// TIA Portal project "kelishangliao" (V15)

(* hardware
DEVICE "S7300/ET200M station_1"  S7-300 station
   slot 0: "导轨_0"  Rail  6ES7 390-1***0-0AA0
   slot 2: "PLC_1"  CPU 314C-2 PN/DP  6ES7 314-6EH04-0AB0  V3.3
      slot 2: "PROFINET 接口_1"  PN-IO
         slot 1: "Port_1"  Port
         slot 2: "Port_2"  Port
      slot 5: "DI 24/DO 16_1"  DI24/DO16
      slot 6: "AI 5/AO 2_1"  AI5/AO2
      slot 7: "计数_1"  Counter
      slot 8: "定位_1"  Positioning
*)

// ===== PLC "PLC_1"  CPU 314C-2 PN/DP =====

VAR_GLOBAL   // PLC tag table "默认变量表"
   "开始按钮" AT %I0.0 : Bool;
   "复位按钮" AT %I0.1 : Bool;
   "停止按钮" AT %I0.4 : Bool;
   "上电" AT %I0.5 : Bool;
   "空瓶到位" AT %I1.0 : Bool;
   "夹瓶处电眼" AT %I1.1 : Bool;
   "颗粒有无" AT %I1.2 : Bool;
   "末端颗粒到位" AT %I1.5 : Bool;
   "主传输带" AT %Q0.0 : Bool;
   "颗粒料传送带" AT %Q0.1 : Bool;
   "旋转气缸" AT %Q0.2 : Bool;
   "升降气缸" AT %Q0.3 : Bool;
   "夹瓶气缸" AT %Q0.4 : Bool;
   "推料颗粒气缸" AT %Q0.5 : Bool;
   "吸盘_电磁阀" AT %Q0.7 : Bool;
   "空瓶输送带_变频器" AT %Q1.0 : Bool;
   "开始灯_绿" AT %Q1.6 : Bool;
   "复位灯_橙" AT %Q1.7 : Bool;
   "M0" AT %M10.0 : Bool;
   "M1" AT %M10.1 : Bool;
   "M2" AT %M10.2 : Bool;
   "M3" AT %M10.3 : Bool;
   "M4" AT %M10.4 : Bool;
   "M5" AT %M10.5 : Bool;
   "M6" AT %M10.6 : Bool;
   "M7" AT %M10.7 : Bool;
   "Tag_1" AT %MD100 : Time;
   "Tag_2" AT %MD104 : Time;
   "Tag_3" AT %MD108 : Time;
   "Tag_4" AT %MD112 : Time;
   "Tag_5" AT %MD116 : Time;
   "Tag_6" AT %MD120 : Time;
   "Tag_7" AT %MD124 : Time;
   "Tag_8" AT %MD128 : Time;
   "Tag_9" AT %MD132 : Time;
   "Tag_10" AT %MW200 : Int;
END_VAR

ORGANIZATION_BLOCK "Main"   // OB1, LAD
TITLE = "Main Program Sweep (Cycle)"
{ S7_Optimized_Access := 'FALSE' }
VERSION : 0.1
   VAR_TEMP
      OB1_EV_CLASS : Byte;   // Bits 0-3 = 1 (Coming event), Bits 4-7 = 1 (Event class 1)
      OB1_SCAN_1 : Byte;   // 1 (Cold restart scan 1 of OB 1), 3 (Scan 2-n of OB 1)
      OB1_PRIORITY : Byte;   // Priority of OB Execution
      OB1_OB_NUMBR : Byte;   // 1 (Organization block 1, OB1)
      OB1_RESERVED_1 : Byte;   // Reserved for system
      OB1_RESERVED_2 : Byte;   // Reserved for system
      OB1_PREV_CYCLE : Int;   // Cycle time of previous OB1 scan (milliseconds)
      OB1_MIN_CYCLE : Int;   // Minimum cycle time of OB1 (milliseconds)
      OB1_MAX_CYCLE : Int;   // Maximum cycle time of OB1 (milliseconds)
      OB1_DATE_TIME : Date_And_Time;   // Date and time OB1 started
   END_VAR
   VAR_TEMP   // added for the SCL form of the ladder/FBD networks
      _w1 : Bool;
   END_VAR
BEGIN

REGION Network 1
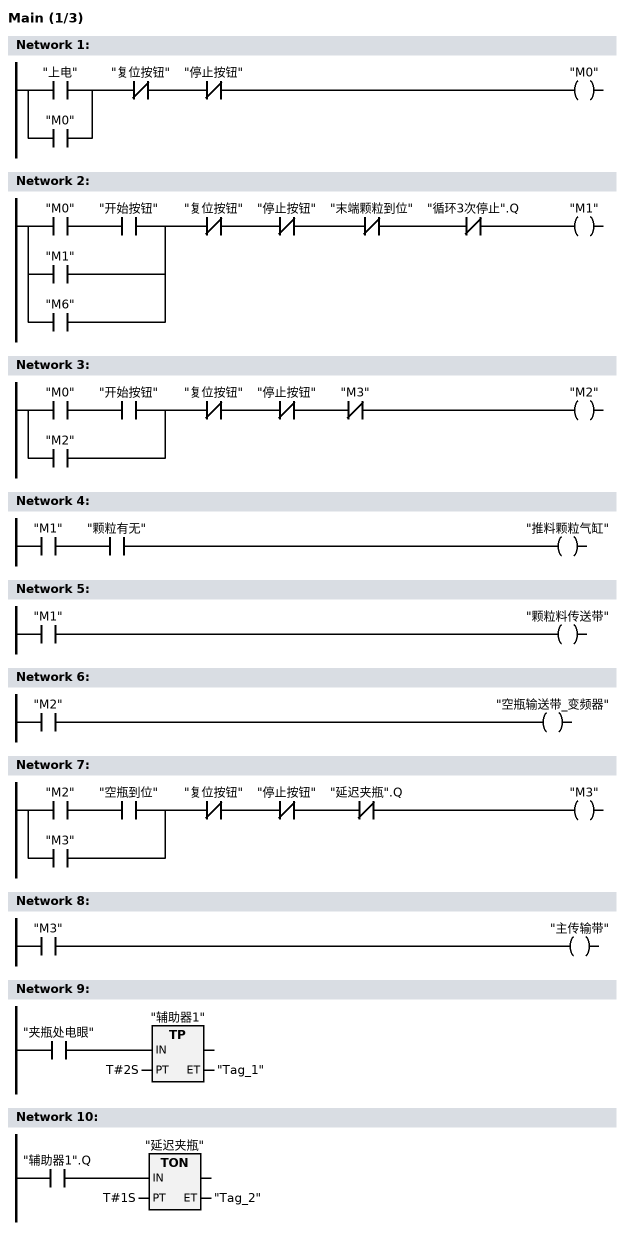
   RUNG wire#powerrail
      Contact( "上电" )
      wire#w1
      I_Contact( "复位按钮" )
      I_Contact( "停止按钮" )
      Coil( "M0" )
   END_RUNG
   RUNG wire#powerrail
      Contact( "M0" )
   END_RUNG wire#w1
   // the same network as SCL:
   "M0" := ("上电" OR "M0") AND NOT "复位按钮" AND NOT "停止按钮";
END_REGION

REGION Network 2
   RUNG wire#powerrail
      Contact( "M0" )
      Contact( "开始按钮" )
      wire#w1
      I_Contact( "复位按钮" )
      I_Contact( "停止按钮" )
      I_Contact( "末端颗粒到位" )
      I_Contact( "循环3次停止".Q )
      Coil( "M1" )
   END_RUNG
   RUNG wire#powerrail
      Contact( "M1" )
   END_RUNG wire#w1
   RUNG wire#powerrail
      Contact( "M6" )
   END_RUNG wire#w1
   // the same network as SCL:
   "M1" := (("M0" AND "开始按钮") OR "M1" OR "M6") AND NOT "复位按钮" AND NOT "停止按钮" AND NOT "末端颗粒到位" AND NOT "循环3次停止".Q;
END_REGION

REGION Network 3
   RUNG wire#powerrail
      Contact( "M0" )
      Contact( "开始按钮" )
      wire#w1
      I_Contact( "复位按钮" )
      I_Contact( "停止按钮" )
      I_Contact( "M3" )
      Coil( "M2" )
   END_RUNG
   RUNG wire#powerrail
      Contact( "M2" )
   END_RUNG wire#w1
   // the same network as SCL:
   "M2" := (("M0" AND "开始按钮") OR "M2") AND NOT "复位按钮" AND NOT "停止按钮" AND NOT "M3";
END_REGION

REGION Network 4
   RUNG wire#powerrail
      Contact( "M1" )
      Contact( "颗粒有无" )
      Coil( "推料颗粒气缸" )
   END_RUNG
   // the same network as SCL:
   "推料颗粒气缸" := "M1" AND "颗粒有无";
END_REGION

REGION Network 5
   RUNG wire#powerrail
      Contact( "M1" )
      Coil( "颗粒料传送带" )
   END_RUNG
   // the same network as SCL:
   "颗粒料传送带" := "M1";
END_REGION

REGION Network 6
   RUNG wire#powerrail
      Contact( "M2" )
      Coil( "空瓶输送带_变频器" )
   END_RUNG
   // the same network as SCL:
   "空瓶输送带_变频器" := "M2";
END_REGION

REGION Network 7
   RUNG wire#powerrail
      Contact( "M2" )
      Contact( "空瓶到位" )
      wire#w1
      I_Contact( "复位按钮" )
      I_Contact( "停止按钮" )
      I_Contact( "延迟夹瓶".Q )
      Coil( "M3" )
   END_RUNG
   RUNG wire#powerrail
      Contact( "M3" )
   END_RUNG wire#w1
   // the same network as SCL:
   "M3" := (("M2" AND "空瓶到位") OR "M3") AND NOT "复位按钮" AND NOT "停止按钮" AND NOT "延迟夹瓶".Q;
END_REGION

REGION Network 8
   RUNG wire#powerrail
      Contact( "M3" )
      Coil( "主传输带" )
   END_RUNG
   // the same network as SCL:
   "主传输带" := "M3";
END_REGION

REGION Network 9
   "辅助器1".TP(IN := "夹瓶处电眼", PT := T#2S, ET => "Tag_1");
END_REGION

REGION Network 10
   "延迟夹瓶".TON(IN := "辅助器1".Q, PT := T#1S, ET => "Tag_2");
END_REGION

REGION Network 11
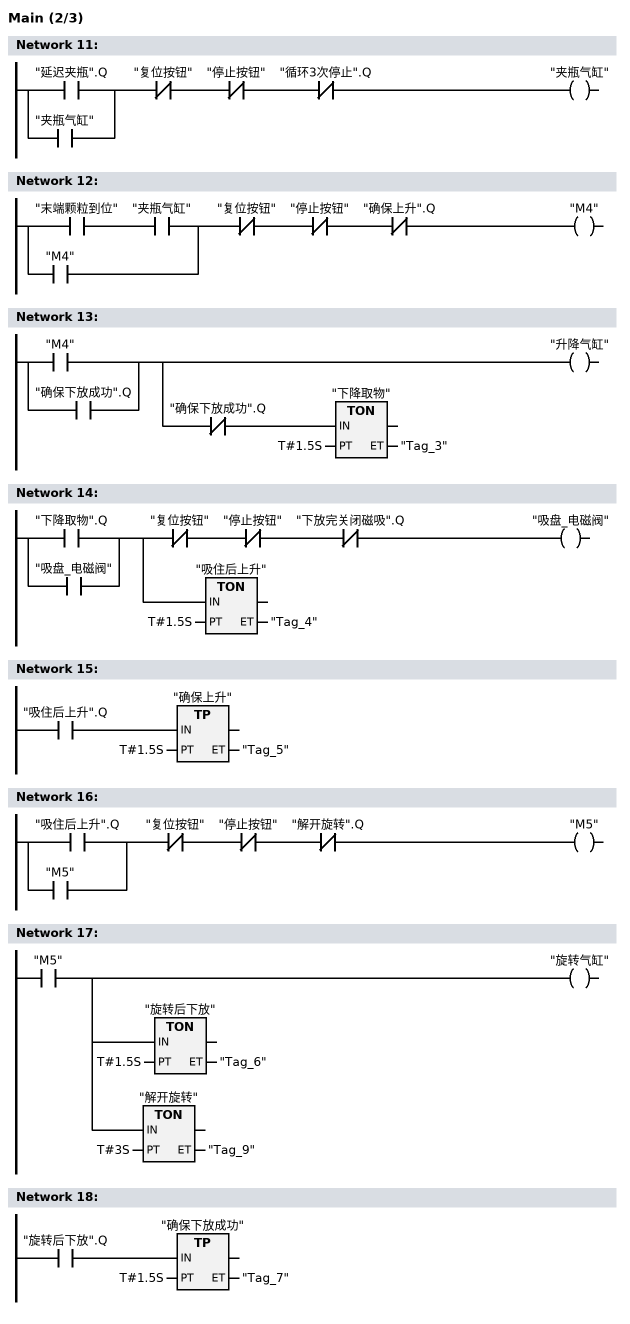
   RUNG wire#powerrail
      Contact( "延迟夹瓶".Q )
      wire#w1
      I_Contact( "复位按钮" )
      I_Contact( "停止按钮" )
      I_Contact( "循环3次停止".Q )
      Coil( "夹瓶气缸" )
   END_RUNG
   RUNG wire#powerrail
      Contact( "夹瓶气缸" )
   END_RUNG wire#w1
   // the same network as SCL:
   "夹瓶气缸" := ("延迟夹瓶".Q OR "夹瓶气缸") AND NOT "复位按钮" AND NOT "停止按钮" AND NOT "循环3次停止".Q;
END_REGION

REGION Network 12
   RUNG wire#powerrail
      Contact( "末端颗粒到位" )
      Contact( "夹瓶气缸" )
      wire#w1
      I_Contact( "复位按钮" )
      I_Contact( "停止按钮" )
      I_Contact( "确保上升".Q )
      Coil( "M4" )
   END_RUNG
   RUNG wire#powerrail
      Contact( "M4" )
   END_RUNG wire#w1
   // the same network as SCL:
   "M4" := (("末端颗粒到位" AND "夹瓶气缸") OR "M4") AND NOT "复位按钮" AND NOT "停止按钮" AND NOT "确保上升".Q;
END_REGION

REGION Network 13
   "升降气缸" := "M4" OR "确保下放成功".Q;
   "下降取物".TON(IN := "升降气缸" AND NOT "确保下放成功".Q, PT := T#1.5S, ET => "Tag_3");
END_REGION

REGION Network 14
   #_w1 := "下降取物".Q OR "吸盘_电磁阀";
   "吸盘_电磁阀" := #_w1 AND NOT "复位按钮" AND NOT "停止按钮" AND NOT "下放完关闭磁吸".Q;
   "吸住后上升".TON(IN := #_w1, PT := T#1.5S, ET => "Tag_4");
END_REGION

REGION Network 15
   "确保上升".TP(IN := "吸住后上升".Q, PT := T#1.5S, ET => "Tag_5");
END_REGION

REGION Network 16
   RUNG wire#powerrail
      Contact( "吸住后上升".Q )
      wire#w1
      I_Contact( "复位按钮" )
      I_Contact( "停止按钮" )
      I_Contact( "解开旋转".Q )
      Coil( "M5" )
   END_RUNG
   RUNG wire#powerrail
      Contact( "M5" )
   END_RUNG wire#w1
   // the same network as SCL:
   "M5" := ("吸住后上升".Q OR "M5") AND NOT "复位按钮" AND NOT "停止按钮" AND NOT "解开旋转".Q;
END_REGION

REGION Network 17
   "旋转气缸" := "M5";
   "旋转后下放".TON(IN := "M5", PT := T#1.5S, ET => "Tag_6");
   "解开旋转".TON(IN := "M5", PT := T#3S, ET => "Tag_9");
END_REGION

REGION Network 18
   "确保下放成功".TP(IN := "旋转后下放".Q, PT := T#1.5S, ET => "Tag_7");
END_REGION

REGION Network 19
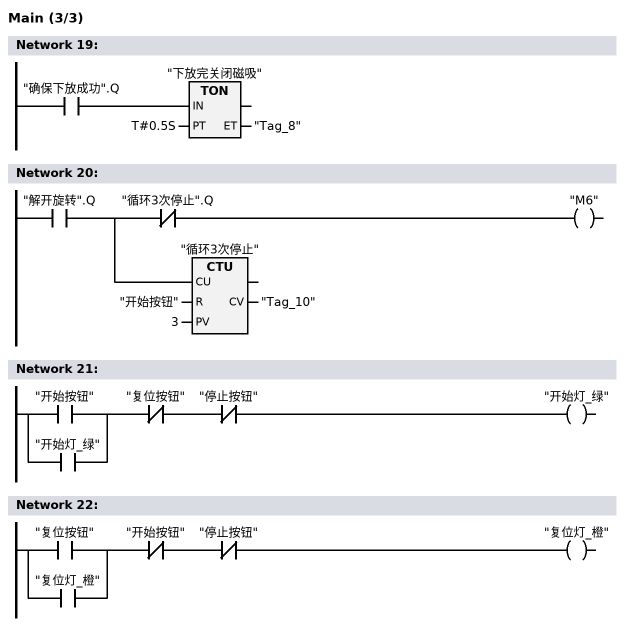
   "下放完关闭磁吸".TON(IN := "确保下放成功".Q, PT := T#0.5S, ET => "Tag_8");
END_REGION

REGION Network 20
   "M6" := "解开旋转".Q AND NOT "循环3次停止".Q;
   "循环3次停止".CTU(CU := "解开旋转".Q, R := "开始按钮", PV := 3, CV => "Tag_10");
END_REGION

REGION Network 21
   RUNG wire#powerrail
      Contact( "开始按钮" )
      wire#w1
      I_Contact( "复位按钮" )
      I_Contact( "停止按钮" )
      Coil( "开始灯_绿" )
   END_RUNG
   RUNG wire#powerrail
      Contact( "开始灯_绿" )
   END_RUNG wire#w1
   // the same network as SCL:
   "开始灯_绿" := ("开始按钮" OR "开始灯_绿") AND NOT "复位按钮" AND NOT "停止按钮";
END_REGION

REGION Network 22
   RUNG wire#powerrail
      Contact( "复位按钮" )
      wire#w1
      I_Contact( "开始按钮" )
      I_Contact( "停止按钮" )
      Coil( "复位灯_橙" )
   END_RUNG
   RUNG wire#powerrail
      Contact( "复位灯_橙" )
   END_RUNG wire#w1
   // the same network as SCL:
   "复位灯_橙" := ("复位按钮" OR "复位灯_橙") AND NOT "开始按钮" AND NOT "停止按钮";
END_REGION
END_ORGANIZATION_BLOCK